Fanuc KAREL source: KO00099.KL

PROGRAM KO00099
%NOLOCKGROUP
VAR
  A: INTEGER
  B: REAL
  OUT: INTEGER
BEGIN
  A = 1
  B = 2
  OUT = ATAN2(A, B)
END KO00099
